(* IEC 61131-3 sources: plc-st-test/test/security/fixtures/injection/src, 1 file *)

(* ---- FB_Dummy.st ---- *)
FUNCTION_BLOCK FB_Dummy
VAR_OUTPUT
  nValue : DINT;
END_VAR
nValue := 1;
END_FUNCTION_BLOCK
